TYPE "ST_CondRecord"
VERSION : 0.1
   STRUCT
      Label : String[120];
      Ok : Bool;
   END_STRUCT;

END_TYPE

